// TIA Portal V20 export
DATA_BLOCK "T4_Resultado"   // DB41901
{ S7_Optimized_Access := 'TRUE' }
AUTHOR : IA
FAMILY : PRUEBA
VERSION : 0.1
// Tanda 1: un Bool por prueba (L_ = KOP, S_ = SCL)
// stored: AutoNumber false
   VAR
      L_I_Coil : Bool;   // Bobina negada -( / )-
      L_SR : Bool;   // Biestable SR (S_SR)
      L_P_Contact : Bool;   // Contacto flanco positivo -|P|-
      L_N_Contact : Bool;   // Contacto flanco negativo -|N|-
      L_NBox : Bool;   // Flanco negativo N_TRIG
      L_P_Coil : Bool;   // Bobina flanco positivo -(P)-
      S_R_TRIG : Bool;   // [SCL] R_TRIG
      S_F_TRIG : Bool;   // [SCL] F_TRIG
      L_TP : Bool;   // Temporizador TP
      L_TOF : Bool;   // Temporizador TOF
      L_TONR : Bool;   // Temporizador TONR
      S_TP : Bool;   // [SCL] TP
      S_TON : Bool;   // [SCL] TON
      S_TOF : Bool;   // [SCL] TOF
      S_TONR : Bool;   // [SCL] TONR
      L_CTU : Bool;   // Contador CTU
      L_CTD : Bool;   // Contador CTD
      L_CTUD : Bool;   // Contador CTUD
      S_CTU : Bool;   // [SCL] CTU
      S_CTD : Bool;   // [SCL] CTD
      S_CTUD : Bool;   // [SCL] CTUD
      L_Mod : Bool;   // Mod (resto)
      S_Mod : Bool;   // [SCL] Mod (resto)
      L_Neg : Bool;   // Neg (cambio de signo)
      S_Neg : Bool;   // [SCL] Neg (cambio de signo)
      L_Abs : Bool;   // Abs (valor absoluto)
      S_Abs : Bool;   // [SCL] Abs (valor absoluto)
      S_Min : Bool;   // [SCL] Min
      S_Max : Bool;   // [SCL] Max
      S_Limit : Bool;   // [SCL] Limit
      L_Sqr : Bool;   // Sqr
      S_Sqr : Bool;   // [SCL] Sqr
      L_Sqrt : Bool;   // Sqrt
      S_Sqrt : Bool;   // [SCL] Sqrt
      L_Ln : Bool;   // Ln
      S_Ln : Bool;   // [SCL] Ln
      L_Exp : Bool;   // Exp
      S_Exp : Bool;   // [SCL] Exp
      L_Sin : Bool;   // Sin
      S_Sin : Bool;   // [SCL] Sin
      L_Cos : Bool;   // Cos
      S_Cos : Bool;   // [SCL] Cos
      L_Tan : Bool;   // Tan
      S_Tan : Bool;   // [SCL] Tan
      L_Frac : Bool;   // Frac
      S_Frac : Bool;   // [SCL] Frac
      L_Asin : Bool;   // Asin
      S_Asin : Bool;   // [SCL] Asin
      L_Acos : Bool;   // Acos
      S_Acos : Bool;   // [SCL] Acos
      L_Atan : Bool;   // Atan
      S_Atan : Bool;   // [SCL] Atan
      S_Expt : Bool;   // [SCL] Expt (potencia)
      S_Inc_Dec : Bool;   // [SCL] INC / DEC no existen en SCL: x := x + 1
      S_MOVE_BLK : Bool;   // [SCL] MOVE_BLK
      S_FILL_BLK : Bool;   // [SCL] FILL_BLK
      S_MOVE_BLK_VARIANT : Bool;   // [SCL] MOVE_BLK_VARIANT
      S_CountOfElements : Bool;   // [SCL] CountOfElements (dentro de una FC con parámetro Variant)
      S_SWAP : Bool;   // [SCL] SWAP
      L_Round : Bool;   // Round
      S_Round : Bool;   // [SCL] Round
      L_Ceil : Bool;   // Ceil
      S_Ceil : Bool;   // [SCL] Ceil
      L_Floor : Bool;   // Floor
      S_Floor : Bool;   // [SCL] Floor
      L_Trunc : Bool;   // Trunc
      S_Trunc : Bool;   // [SCL] Trunc
      S_SCALE_X : Bool;   // [SCL] SCALE_X
      S_NORM_X : Bool;   // [SCL] NORM_X
      L_And : Bool;   // AND
      S_And : Bool;   // [SCL] AND
      L_Or : Bool;   // OR
      S_Or : Bool;   // [SCL] OR
      L_Xor : Bool;   // XOR
      S_Xor : Bool;   // [SCL] XOR
      L_Inv : Bool;   // INV
      S_Inv : Bool;   // [SCL] NOT de Word
      L_Mux : Bool;   // MUX
      L_Demux : Bool;   // DEMUX
      S_Deco : Bool;   // [SCL] DECO
      S_Enco : Bool;   // [SCL] ENCO
      S_Sel : Bool;   // [SCL] SEL
      S_Mux : Bool;   // [SCL] MUX
      L_Shr : Bool;   // SHR
      S_Shr : Bool;   // [SCL] SHR
      L_Shl : Bool;   // SHL
      S_Shl : Bool;   // [SCL] SHL
      L_Ror : Bool;   // ROR
      S_Ror : Bool;   // [SCL] ROR
      L_Rol : Bool;   // ROL
      S_Rol : Bool;   // [SCL] ROL
      S_REPEAT : Bool;   // [SCL] REPEAT / UNTIL
      S_EXIT_CONTINUE : Bool;   // [SCL] EXIT y CONTINUE
      S_GOTO : Bool;   // [SCL] GOTO y etiqueta
      S_RUNTIME : Bool;   // [SCL] RUNTIME
      S_GET_ERR_ID : Bool;   // [SCL] GET_ERR_ID
      Vida : DInt;   // Sube cada ciclo si T4_Base se ejecuta
      OK : Int;   // Pruebas correctas
      Total : Int := 96;   // Pruebas
      Todo_OK : Bool;   // Todas correctas
   END_VAR
BEGIN
END_DATA_BLOCK
